Staubli VAL3: Lab2B_Level2.pjx

--- Lab2B_Level2.pjx ---
parameters version=s6.8 stackSize=5000 millimeterUnit=true
program file=start.pgx
program file=feedCylinder.pgx
program file=assemble.pgx
program file=placeAssembly.pgx
program file=physicalIO.pgx
program file=stop.pgx
data file=Lab2B_Level2.dtx
alias name=io interface=io autoload=true

--- Lab2B_Level2.dtx ---


--- start.pgx ---
program start()
// Level 2 - four assemblies; validate setup and trajectories in SRS.
  local num poseIndex
  local point approachPose
  local point placePose
begin
  // ============================================================
  // LEVEL 2: ALIMENTAR, MONTAR Y COLOCAR CUATRO CONJUNTOS
  // ============================================================
  // Aplicacion separada: Lab2B (Level 1) permanece sin modificar.
  // Matriz VACIA y cuatro pistones cargados al comenzar.
  // simulation=true: sensores manuales, sin acceso a pines.
  // simulation=false: bIn2/14/15, bOut10 y pinza valve1.
  userPage()
  cls()
  putln("Lab2B_Level2 - Four assemblies - empty matrix required")
  physicalRun = !simulation
  placedCount = 0
  partIndex = 0
  cycleStep = 0
  feederExtend = false
  ioReady = false

  // ============================================================
  // COMPROBAR ALTURAS DE MATRIZ SIN MOVER NI ACCIONAR SALIDAS
  // ============================================================
  // Parejas 0/1, 2/3, 4/5, 6/7: par=approach, impar=deposito.
  // J3 es un ANGULO, no una altura. Calculamos Z del TCP lateral.
  // Esto comprueba altura, no colisiones, alineacion o alcance del trayecto.
  for poseIndex = 0 to 3
    approachPose = jointToPoint(tLateral, world, jMatrix[2*poseIndex])
    placePose = jointToPoint(tLateral, world, jMatrix[2*poseIndex+1])
    putln("Matrix slot (0..3):")
    putln(poseIndex)
    putln("Approach Z (mm):")
    putln(approachPose.trsf.z)
    putln("Place Z (mm):")
    putln(placePose.trsf.z)
    if approachPose.trsf.z <= placePose.trsf.z
      putln("ERROR: approach is not above place; review this matrix pair")
      return
    endIf
  endFor

  // ============================================================
  // LOS CUATRO PISTONES TODAVIA ESTAN POR ENSENAR
  // ============================================================
  // jPistonPick[0..7] esta a cero a proposito. No reutilizamos
  // cuatro veces la unica recogida del Level 1 ni inventamos offsets.
  // Completar las OCHO posturas: par=approach, impar=recogida.
  // Este control termina ANTES de crear tareas o dar ordenes al robot.
  for poseIndex = 0 to 7
    if jPistonPick[poseIndex].j1 == 0 and jPistonPick[poseIndex].j2 == 0 and jPistonPick[poseIndex].j3 == 0 and jPistonPick[poseIndex].j4 == 0 and jPistonPick[poseIndex].j5 == 0 and jPistonPick[poseIndex].j6 == 0
      putln("ERROR: teach piston approach/pick joint; missing index:")
      putln(poseIndex)
      return
    endIf
  endFor

  // physicalIO solo escribe el ALIMENTADOR; nunca la pinza.
  if physicalRun
    taskCreate "physicalIO", 10, physicalIO()
    wait(ioReady == true)
    putln("PHYSICAL: real sensors and feeder enabled")
    open(tLateral)
  else
    putln("MANUAL SIMULATION: change sensor bools at the indicated steps")
    delay(tLateral.otime)
  endIf
  movej(jStart[0], tLateral, mNomSpeed)
  waitEndMove()

  // ============================================================
  // SOLO CUATRO CONJUNTOS; NO HAY QUINTA ALIMENTACION
  // ============================================================
  while placedCount < 4
    partIndex = placedCount
    putln("Assembly number (1..4):")
    putln(partIndex+1)
    call feedCylinder()
    call assemble()
    call placeAssembly()
    // Contar tras soltar y terminar la retirada de la matriz.
    placedCount = placedCount + 1
    putln("Completed matrix slots:")
    putln(placedCount)
    // Volver a la postura inicial SOLO si falta otro conjunto.
    if placedCount < 4
      movej(jStart[0], tLateral, mNomSpeed)
      waitEndMove()
    endIf
  endWhile

  // La matriz llena finaliza aunque bIn2 siga detectando cilindros.
  feederExtend = false
  taskKill("physicalIO")
  if physicalRun
    io:bOut10 = false
  endIf
  ioReady = false
  cycleStep = 100
  putln("100 - Matrix full: 4/4. No further feeding or pickup.")
end

--- assemble.pgx ---
program assemble()
// Level 2 - four assemblies; validate setup and trajectories in SRS.
begin
  // partIndex=0..3 selecciona la pareja del piston correspondiente.
  // ============================================================
  // 20. RECOGER EL CILINDRO CON EL TCP LATERAL
  // ============================================================
  // movej: traslado articular entre aproximaciones.
  // movel: entradas/retiradas con mApproachSpeed; insercion con mInsertSpeed.
  // jointToPoint convierte la joint para movel; no mueve el robot.
  // Usar el mismo TCP en la conversion y en la orden de movimiento.
  // waitEndMove termina cada movimiento antes de accionar la pinza.
  cycleStep = 20
  putln("20 - Pick cylinder - tLateral")
  movej(jCylinderPick[0], tLateral, mNomSpeed)
  waitEndMove()
  movel(jointToPoint(tLateral, world, jCylinderPick[1]), tLateral, mApproachSpeed)
  waitEndMove()

  // Cerrar y dar el tiempo mecanico guardado en la herramienta (1 s).
  // No hay confirmacion de agarre en el mapa de E/S de esta practica.
  if physicalRun
    close(tLateral)
  else
    delay(tLateral.ctime)
  endIf
  movel(jointToPoint(tLateral, world, jCylinderPick[0]), tLateral, mApproachSpeed)
  waitEndMove()
  // El cilindro ya se ha retirado: exigir sensor libre antes
  // de admitir otra alimentacion en la siguiente vuelta.
  cycleStep = 21
  putln("21 - Wait cylinderPresent=false after cylinder withdrawal")
  wait(cylinderPresent == false)

  // ============================================================
  // 30. DEPOSITAR EL CILINDRO EN LA ESTACION DE MONTAJE
  // ============================================================
  cycleStep = 30
  putln("30 - Place cylinder at assembly station")
  movej(jCylinderPlace[0], tLateral, mNomSpeed)
  waitEndMove()
  movel(jointToPoint(tLateral, world, jCylinderPlace[1]), tLateral, mApproachSpeed)
  waitEndMove()
  if physicalRun
    open(tLateral)
  else
    delay(tLateral.otime)
  endIf
  movel(jointToPoint(tLateral, world, jCylinderPlace[0]), tLateral, mApproachSpeed)
  waitEndMove()

  // ============================================================
  // 40. RECOGER EL PISTON CON EL TCP DE PUNTA
  // ============================================================
  // tTip y tLateral son DOS TCP de LA MISMA PINZA y salida valve1.
  // Cambiar de TCP no cambia fisicamente la herramienta.
  // Level 1 supone un piston en el punto ensenado; no espera bIn0.
  cycleStep = 40
  putln("40 - Pick piston - tTip")
  if physicalRun
    open(tTip)
  else
    delay(tTip.otime)
  endIf
  putln("DBG 40A - BEFORE movej: selected piston approach")
  movej(jPistonPick[2*partIndex], tTip, mNomSpeed)
  waitEndMove()
  putln("DBG 40B - Approach reached; BEFORE movel: selected piston pick")
  movel(jointToPoint(tTip, world, jPistonPick[2*partIndex+1]), tTip, mApproachSpeed)
  waitEndMove()
  putln("DBG 40C - Pick reached; sending CLOSE command")
  if physicalRun
    close(tTip)
  else
    delay(tTip.ctime)
  endIf
  putln("DBG 40D - close(tTip) completed; closing time included")
  // Diagnostico despues de close(tTip), que ya incluye ctime.
  // El adaptador no escribe la pinza; solo lee el sensor de cilindro.
  putln("DBG 40E - Closing delay finished; cycleStep:")
  putln(cycleStep)
  putln("DBG Last gripper command: close(tTip)")
  if physicalRun
    putln("DBG physicalRun=true; physicalIO task status:")
    putln(taskStatus("physicalIO"))
    putln("DBG task status: 1=running, 0=suspended, -1=absent, other=error")
    if ioReady and taskStatus("physicalIO") == 1
      if io:valve1 == true
        putln("DBG valve1=1 (OPEN output)")
      else
        putln("DBG valve1=0 (CLOSE output)")
      endIf
    else
      putln("DBG valve1 not read: IO task not ready/running")
    endIf
  else
    putln("DBG physicalRun=false; manual simulation, no pin access")
  endIf
  putln("DBG 40F - BEFORE movel: withdraw to selected piston approach")
  movel(jointToPoint(tTip, world, jPistonPick[2*partIndex]), tTip, mApproachSpeed)
  waitEndMove()
  putln("DBG 40G - Withdrawal completed; leaving piston pickup")

  // ============================================================
  // 50. INSERTAR EL PISTON Y SOLTARLO ANTES DE RETIRARSE
  // ============================================================
  // TODO SIMULACION: confirmar el orden [0]/[1] de gridpiston.
  // TODO FISICO: ajustar alineacion y profundidad de jPistonInsert[1].
  // Este movimiento es por posicion; no mide fuerza ni confirma montaje.
  cycleStep = 50
  putln("50 - Insert piston into cylinder")
  putln("DBG 50A - BEFORE movej: insertion approach [0]")
  movej(jPistonInsert[0], tTip, mNomSpeed)
  waitEndMove()
  putln("DBG 50B - Insertion approach reached")
  movel(jointToPoint(tTip, world, jPistonInsert[1]), tTip, mInsertSpeed)
  waitEndMove()
  putln("DBG 50C - Insertion reached with tTip; opening gripper")
  if physicalRun
    open(tTip)
  else
    delay(tTip.otime)
  endIf
  putln("DBG 50D - BEFORE withdrawal with tTip to jPistonInsert[0]")
  movel(jointToPoint(tTip, world, jPistonInsert[0]), tTip, mInsertSpeed)
  waitEndMove()
  putln("DBG 50E - Tip withdrawal completed")

  // ============================================================
  // 55. POSTURA INTERMEDIA ANTES DE RECOGER EL CONJUNTO
  // ============================================================
  // Joint indicada por el usuario. Se alcanza DESPUES de soltar
  // el piston y retirarse con tTip, antes del agarre con tLateral.
  cycleStep = 55
  putln("DBG 55A - BEFORE movej: jAssemblyMove with tTip")
  movej(jAssemblyMove, tTip, mNomSpeed)
  waitEndMove()
  putln("DBG 55B - Assembly transit posture reached")

end

--- feedCylinder.pgx ---
program feedCylinder()
// Level 2 - four assemblies; validate setup and trajectories in SRS.
begin
  // ============================================================
  // PREPARAR UN CILINDRO, CON EL ROBOT FUERA DEL DISPENSADOR
  // ============================================================
  // bOut10: 1=extender, 0=retraer (mapa del enunciado).
  // bIn14/bIn15: finales extendido/retraido; bIn2: cilindro listo.
  // El PDF no especifica toda la secuencia mecanica: se propone
  // extender y retraer antes de entrar con el robot. Verificar en la celda.
  // Si ya hay un cilindro preparado, no empujar otro encima.
  cycleStep = 10
  feederExtend = false
  putln("10 - Wait feederRetracted=true and feederExtended=false")
  wait(feederRetracted == true and feederExtended == false)
  if !cylinderPresent
    cycleStep = 11
    putln("11 - EXTEND feeder; wait extended=true / retracted=false")
    feederExtend = true
    wait(feederExtended == true and feederRetracted == false)

    cycleStep = 12
    putln("12 - RETRACT feeder; wait retracted=true / extended=false")
    feederExtend = false
    wait(feederRetracted == true and feederExtended == false)
  endIf
  cycleStep = 13
  putln("13 - Wait cylinderPresent=true; cylinder ready for pickup")
  wait(cylinderPresent == true)
end

--- physicalIO.pgx ---
program physicalIO()
// Level 2 - four assemblies; validate setup and trajectories in SRS.
begin
  // ============================================================
  // SENSORES Y ALIMENTADOR DEL LEVEL 2
  // ============================================================
  // Solo se crea en fisico. En simulacion los sensores se editan a mano.
  // La pinza usa open/close con valve1; NO escribir valve1 aqui.
  while true
    cylinderPresent = io:bIn2 == true
    feederExtended = io:bIn14 == true
    feederRetracted = io:bIn15 == true
    io:bOut10 = feederExtend
    ioReady = true
    delay(0.01)
  endWhile
end

--- placeAssembly.pgx ---
program placeAssembly()
// Level 2 - four assemblies; validate setup and trajectories in SRS.
begin
  // ============================================================
  // 60. RECOGER EL CONJUNTO CON EL TCP LATERAL
  // ============================================================
  // Recoger en jCylinderPlace[1], donde se ha depositado el cilindro.
  // TODO FISICO: comprobar el agarre con el piston ya dentro del cilindro.
  cycleStep = 60
  putln("60 - Pick assembled cylinder - tLateral")
  if physicalRun
    open(tLateral)
  else
    delay(tLateral.otime)
  endIf
  // El siguiente movimiento usa el TCP lateral. Las joints guardadas
  // deben describir la postura de agarre lateral; el TCP no anade un giro.
  putln("DBG 60A - BEFORE movej with tLateral to jCylinderPlace[0]")
  movej(jCylinderPlace[0], tLateral, mNomSpeed)
  waitEndMove()
  putln("DBG 60B - Lateral approach reached; BEFORE descent to jCylinderPlace[1]")
  movel(jointToPoint(tLateral, world, jCylinderPlace[1]), tLateral, mApproachSpeed)
  waitEndMove()
  putln("DBG 60C - Assembly pickup reached with tLateral; closing gripper")
  if physicalRun
    close(tLateral)
  else
    delay(tLateral.ctime)
  endIf
  putln("DBG 60D - BEFORE withdrawal of assembly with tLateral")
  movel(jointToPoint(tLateral, world, jCylinderPlace[0]), tLateral, mApproachSpeed)
  waitEndMove()
  putln("DBG 60E - Assembly withdrawal completed")

  // ============================================================
  // DEPOSITAR EN LA PAREJA DEL HUECO ACTUAL DE LA MATRIZ
  // ============================================================
  // partIndex es 0..3: approach=2*i, deposito=2*i+1.
  cycleStep = 70
  putln("70 - Place assembly in matrix slot (0..3):")
  putln(partIndex)
  movej(jMatrix[2*partIndex], tLateral, mNomSpeed)
  waitEndMove()
  movel(jointToPoint(tLateral, world, jMatrix[2*partIndex+1]), tLateral, mApproachSpeed)
  waitEndMove()
  if physicalRun
    open(tLateral)
  else
    delay(tLateral.otime)
  endIf
  movel(jointToPoint(tLateral, world, jMatrix[2*partIndex]), tLateral, mApproachSpeed)
  waitEndMove()
  putln("75 - Assembly released; matrix withdrawal completed")
end

--- stop.pgx ---
program stop()
// Level 2 - four assemblies; validate setup and trajectories in SRS.
begin
  // Detener el adaptador antes de mandar retraer el alimentador.
  // taskKill no hace nada si la tarea no existe (p. ej. setup incompleto).
  taskKill("physicalIO")
  resetMotion()
  feederExtend = false
  // No tocar hardware si start termino por posiciones pendientes.
  if physicalRun and ioReady
    io:bOut10 = false
  endIf
  ioReady = false
  cycleStep = -1
  // No abrir/cerrar la pinza ni ordenar retorno automatico.
  // Un nuevo start reinicia el contador: vaciar matriz antes de reiniciar.
  putln("STOP - Feeder retract command; gripper unchanged. Prepare cell before restart.")
end
